    rq_activate_all_grippers(True)
    # end: URCap Program Node
  end
  $ 55 "zero_ftsensor()"
  zero_ftsensor()
  $ 56 "EXTT"
  $ 57 "Set GRP_3F_Enable=Off"
  set_standard_digital_out(4, False)
  $ 58 "Set BarcodeTrigger=Off"
  set_standard_digital_out(6, False)
  $ 59 "Set GRP_3F_Decap=Off"
  set_standard_digital_out(3, False)
  $ 60 "Set GRP_3F_Cap=Off"
  set_standard_digital_out(2, False)
  $ 61 "Set GRP_3F_Open=Off"
  set_standard_digital_out(5, False)
  $ 62 "PSE_T≔get_tool_free_pose(dir=[0,0,0.150], move_in_base_frame=True)"
  global PSE_T=get_tool_free_pose(dir=[0,0,0.150], move_in_base_frame=True)
  $ 63 "If is_reachable(Base_const, [PSE_T])"
  if (is_reachable(p[0.0,0.0,0.0,0.0,0.0,0.0], [PSE_T])):
    $ 64 "MoveL"
    $ 65 "PSE_T" "breakAfter"
    movel(PSE_T, a=1.2, v=0.15)
  end
  while (True):
    $ 66 "Robot Program"
    $ 67 "MAIN"
    $ 68 "command_manager(external_control='uGO', cond_suspend=(ITM_Manipulated and AMR_AtTarget and AMR_Charging and AMR_Battery<40), cond_unsuspend=(AMR_Battery≟60))"
    command_manager(external_control="uGO", cond_suspend=(ITM_Manipulated  and  AMR_AtTarget  and  AMR_Charging  and  AMR_Battery<40), cond_unsuspend=(AMR_Battery == 60))
    $ 69 "log_state(STATE_Info)"
    log_state(STATE_Info)
    $ 70 "Switch STATE"
    switch_1 = STATE
    $ 71 "Case 1"
    if (1 == switch_1):
      $ 72 "Stopping"
      $ 73 "STATE_Info≔'Stopping'"
      global STATE_Info="Stopping"
      $ 74 "end_freedrive_mode()"
      end_freedrive_mode()
      $ 75 "Set"
      set_tcp(p[0.0,0.0,0.161,3.1415,0.0,0.0])
      $ 76 "PSE_T≔get_tool_free_pose(dir=[0,0,0.150], move_in_base_frame=True)"
      global PSE_T=get_tool_free_pose(dir=[0,0,0.150], move_in_base_frame=True)
      $ 77 "If is_reachable(Base_const, [PSE_T])"
      if (is_reachable(p[0.0,0.0,0.0,0.0,0.0,0.0], [PSE_T])):
        $ 78 "MoveL"
        $ 79 "PSE_T" "breakAfter"
        movel(PSE_T, a=1.2, v=0.15)
      end
      $ 80 "do_transition(keep_rxry=OBJ_Picked, r=0)"
      do_transition(keep_rxry=OBJ_Picked, r=0)
      $ 81 "Decapper"
      $ 82 "Set GRP_3F_Enable=Off"
      set_standard_digital_out(4, False)
      $ 83 "Set BarcodeTrigger=Off"
      set_standard_digital_out(6, False)
      $ 84 "Set GRP_3F_Decap=Off"
      set_standard_digital_out(3, False)
      $ 85 "Set GRP_3F_Cap=Off"
      set_standard_digital_out(2, False)
      $ 86 "Set GRP_3F_Open=Off"
      set_standard_digital_out(5, False)
      $ 89 "Call Sub_AMR_MiR_V3"
      Sub_AMR_MiR_V3()
      $ 90 "If stopping() and AMR_Done"
      if (stopping()  and  AMR_Done):
        $ 91 "STATE≔2"
        global STATE=2
        $ 92 "ugo_update_outputs()"
        ugo_update_outputs()
      end
    elif (2 == switch_1):
      $ 93 "Case 2"
      $ 94 "Stopped"
      $ 95 "STATE_Info≔'Stopped'"
      global STATE_Info="Stopped"
      $ 96 "Call Sub_AMR_MiR_V3"
      Sub_AMR_MiR_V3()
      $ 97 "If CMD_Reset"
      if (CMD_Reset):
        $ 98 "STATE≔3"
        global STATE=3
        $ 99 "ugo_update_outputs()"
        ugo_update_outputs()
      end
    elif (3 == switch_1):
      $ 100 "Case 3"
      $ 101 " Resetting"
      $ 102 "STATE_Info≔'Resetting'"
      global STATE_Info="Resetting"
      $ 103 "uML"
      $ 104 "reset_error()"
      reset_error()
      $ 105 "reset_warning()"
      reset_warning()
      $ 106 "PROCESS_Step≔0"
      global PROCESS_Step=0
      $ 107 "PROCESS_Info≔''"
      global PROCESS_Info=""
      $ 108 "ARM_Referenced≔ False "
      global ARM_Referenced=  False
      $ 109 "WRK_Done≔ False "
      global WRK_Done=  False
      $ 110 "ITM_Prepared≔ False "
      global ITM_Prepared=  False
      $ 111 "ITM_Manipulated≔ False "
      global ITM_Manipulated=  False
      $ 112 "STP≔0"
      global STP=0
      $ 113 "Action≔0"
      global Action=0
      $ 114 "Action_Info≔''"
      global Action_Info=""
      $ 115 "ITM_ID≔0"
      global ITM_ID=0
      $ 116 "JIG≔0"
      global JIG=0
      $ 117 "JIG_Slot≔0"
      global JIG_Slot=0
      $ 118 "Task_info≔''"
      global Task_info=""
      $ 119 "Set"
      set_tcp(p[0.0,0.0,0.161,3.1415,0.0,0.0])
      $ 120 "App"
      $ 121 "'ADD APPLICATION SPECIFIC COMMANDS'"
      # 'ADD APPLICATION SPECIFIC COMMANDS'
      $ 122 "OBJ_Type≔0"
      global OBJ_Type=0
      $ 123 "OBJ_Nbr≔0"
      global OBJ_Nbr=0
      $ 124 "If CNT_Rack_Output≥50"
      if (CNT_Rack_Output >= 50):
        $ 125 "CNT_Rack_Output≔0"
        global CNT_Rack_Output=0
      end
      $ 126 "TASK≔struct(ID=0, NAVI=struct(target=0, footprint=0, protectiveOff=0, dock=0), WORK=struct(ITM_ID_Src=0, JIG_ID_Src=0, OBJ_Nbr_Src=0, ACT_Src=0, ITM_ID_Tgt=0, JIG_ID_Tgt=0, OBJ_Nbr_Tgt=0, ACT_Tgt=0, OBJ_Type=0))"
      global TASK=struct(ID=0, NAVI=struct(target=0, footprint=0, protectiveOff=0, dock=0), WORK=struct(ITM_ID_Src=0, JIG_ID_Src=0, OBJ_Nbr_Src=0, ACT_Src=0, ITM_ID_Tgt=0, JIG_ID_Tgt=0, OBJ_Nbr_Tgt=0, ACT_Tgt=0, OBJ_Type=0))
      $ 127 "Call Sub_AMR_MiR_V3"
      Sub_AMR_MiR_V3()
      $ 128 "If resetting() and AMR_Done"
      if (resetting()  and  AMR_Done):
        $ 129 "STATE≔4"
        global STATE=4
        $ 130 "ugo_update_outputs()"
        ugo_update_outputs()
      end
    elif (4 == switch_1):
      $ 131 "Case 4"
      $ 132 "Idle"
      $ 133 "STATE_Info≔'Idle'"
      global STATE_Info="Idle"
      $ 134 "If CMD_Start"
      if (CMD_Start):
        $ 135 "STATE≔5"
        global STATE=5
        $ 136 "ugo_update_outputs()"
        ugo_update_outputs()
      end
    elif (5 == switch_1):
      $ 137 "Case 5"
      $ 138 "Starting"
      $ 139 "STATE_Info≔'Starting'"
      global STATE_Info="Starting"
      $ 140 "'ADD COMMANDS WHAT TO START WITH'"
      # 'ADD COMMANDS WHAT TO START WITH'
      $ 141 "Call Sub_AMR_MiR_V3"
      Sub_AMR_MiR_V3()
      $ 142 "get ugo data"
      $ 143 "Assign Tasks"
      $ 144 "TASK.ID = ugo_get_task()"
      TASK.ID = ugo_get_task()
      $ 145 "If TASK.ID≟1"
      if (TASK.ID == 1):
        $ 146 "Task_info≔'Charge'"
        global Task_info="Charge"
        $ 147 "Parameters"
        $ 148 "AMR_PosTarget≔1"
        global AMR_PosTarget=1
      else:
        $ 149 "ElseIf TASK.ID≟9"
        if (TASK.ID == 9):
          $ 150 "'Pick Sarstedt Rack from Variable source'"
          # 'Pick Sarstedt Rack from Variable source'
          $ 151 "Task_info≔'Navigate to Target'"
          global Task_info="Navigate to Target"
          $ 152 "Parameters"
          $ 153 "AMR_PosTarget≔UGO.read_input('00','ITM_ID')"
          global AMR_PosTarget=UGO.read_input("00","ITM_ID")
        else:
          $ 154 "ElseIf TASK.ID≟10"
          if (TASK.ID == 10):
            $ 155 "'Pick Sarstedt Rack from Variable source'"
            # 'Pick Sarstedt Rack from Variable source'
            $ 156 "Task_info≔'Pick Rack'"
            global Task_info="Pick Rack"
            $ 157 "AMR_PosTarget≔2"
            global AMR_PosTarget=2
            $ 158 "Parameters"
            $ 159 "ITM_ID≔UGO.read_input('00','ITM_ID')"
            global ITM_ID=UGO.read_input("00","ITM_ID")
            $ 160 "JIG≔UGO.read_input('00','JIG_ID')"
            global JIG=UGO.read_input("00","JIG_ID")
            $ 161 "OBJ_Type≔3"
            global OBJ_Type=3
          else:
            $ 163 "ElseIf TASK.ID≟11"
            if (TASK.ID == 11):
              $ 164 "'Place Sarstedt Rack on Variable target'"
              # 'Place Sarstedt Rack on Variable target'
              $ 165 "Task_info≔'Place Rack'"
              global Task_info="Place Rack"
              $ 166 "AMR_PosTarget≔2"
              global AMR_PosTarget=2
              $ 167 "Parameters"
              $ 168 "ITM_ID≔UGO.read_input('00','ITM_ID')"
              global ITM_ID=UGO.read_input("00","ITM_ID")
              $ 169 "JIG≔UGO.read_input('00','JIG_ID')"
              global JIG=UGO.read_input("00","JIG_ID")
              $ 170 "OBJ_Type≔3"
              global OBJ_Type=3
            else:
              $ 172 "ElseIf TASK.ID≟12"
              if (TASK.ID == 12):
                $ 173 "Task_info≔'Decapping'"
                global Task_info="Decapping"
                $ 174 "Parameters"
                $ 175 "ITM_ID≔1"
                global ITM_ID=1
                $ 176 "AMR_PosTarget≔AMR_PosActual"
                global AMR_PosTarget=AMR_PosActual
                $ 177 "PRC_TubCounter≔0"
                global PRC_TubCounter=0
              else:
                $ 178 "ElseIf TASK.ID≟13"
                if (TASK.ID == 13):
                  $ 179 "Task_info≔'Empty racks'"
                  global Task_info="Empty racks"
                  $ 180 "Parameters"
                  $ 181 "ITM_ID≔1"
                  global ITM_ID=1
                  $ 182 "AMR_PosTarget≔AMR_PosActual"
                  global AMR_PosTarget=AMR_PosActual
                else:
                  $ 183 "ElseIf TASK.ID≟14"
                  if (TASK.ID == 14):
                    $ 184 "Task_info≔'Decap'"
                    global Task_info="Decap"
                    $ 185 "Parameters"
                    $ 186 "ITM_ID≔1"
                    global ITM_ID=1
                    $ 187 "OBJ_Type≔2"
                    global OBJ_Type=2
                    $ 188 "JIG≔7"
                    global JIG=7
                    $ 189 "AMR_PosTarget≔AMR_PosActual"
                    global AMR_PosTarget=AMR_PosActual
                  else:
                    $ 190 "ElseIf TASK.ID≟99"
                    if (TASK.ID == 99):
                      $ 191 "Task_info≔'Decapping and barcode alignment'"
                      global Task_info="Decapping and barcode alignment"
                      $ 192 "Parameters"
                      $ 193 "PRC_TubNumber≔UGO.read_input('00','TubesNb')"
                      global PRC_TubNumber=UGO.read_input("00","TubesNb")
                      $ 194 "PRC_TubCounter≔0"
                      global PRC_TubCounter=0
                      $ 195 "ITM_ID≔1"
                      global ITM_ID=1
                      $ 196 "AMR_PosTarget≔AMR_PosActual"
                      global AMR_PosTarget=AMR_PosActual
                    else:
                      $ 205 "ElseIf TASK.ID≟15"
                      if (TASK.ID == 15):
                        $ 206 "Task_info≔'Unoad Centrifuge'"
                        global Task_info="Unoad Centrifuge"
                        $ 207 "Parameters"
                        $ 208 "PRC_RackCounter≔0"
                        global PRC_RackCounter=0
                        $ 209 "TASK.WORK.ITM_ID_Src=2"
                        TASK.WORK.ITM_ID_Src=2
                        $ 210 "TASK.WORK.ITM_ID_Tgt=1"
                        TASK.WORK.ITM_ID_Tgt=1
                        $ 211 "AMR_PosTarget≔4"
                        global AMR_PosTarget=4
                        $ 212 "AMR_FootprintID≔1"
                        global AMR_FootprintID=1
                      else:
                        $ 231 "Else" "noBreak"
                        $ 232 "set_error(ERROR_WRONG_ORDER)"
                        set_error(ERROR_WRONG_ORDER)
                      end
                    end
                  end
                end
              end
            end
          end
        end
      end
      $ 233 "test ugo"
      $ 234 "Wait: 0.2"
      sleep(0.2)
      $ 235 "ugo_update_outputs()"
      ugo_update_outputs()
      $ 236 "If starting() and AMR_Done"
      if (starting()  and  AMR_Done):
        $ 237 "log_message(Task_info, 'New Task: ')"
        log_message(Task_info, "New Task: ")
        $ 238 "log_message(to_str(TASK.ID), 'Task_ID: ')"
        log_message(to_str(TASK.ID), "Task_ID: ")
        $ 239 "do_transition(keep_rxry=OBJ_Picked)"
        do_transition(keep_rxry=OBJ_Picked)
        $ 240 "STATE≔6"
        global STATE=6
        $ 241 "ugo_update_outputs()"
        ugo_update_outputs()
      end
    elif (6 == switch_1):
      $ 242 "Case 6"
      $ 243 "Execute"
      $ 244 "STATE_Info≔'Execute'"
      global STATE_Info="Execute"
      $ 245 "If  not CMD_Hold and not CMD_Suspend"
      global thread_flag_245=0
      thread Thread_if_245():
        $ 246 "Switch PROCESS_Step"
        switch_2 = PROCESS_Step
        $ 247 "Case 0"
        if (0 == switch_2):
          $ 248 "PROCESS_Info≔'process control'"
          global PROCESS_Info="process control"
          $ 249 "log_process(PROCESS_Info)"
          log_process(PROCESS_Info)
          $ 250 "process control"
          $ 251 "If  not AMR_AtTarget"
          if (  not  AMR_AtTarget):
            $ 252 "PROCESS_Step≔1"
            global PROCESS_Step=1
          else:
            $ 253 "ElseIf (( not ITM_Prepared and  not WRK_Done) or (ITM_Prepared and WRK_Done))"
            if (((  not  ITM_Prepared  and    not  WRK_Done)  or  (ITM_Prepared  and  WRK_Done))):
              $ 254 "PROCESS_Step≔2"
              global PROCESS_Step=2
            else:
              $ 255 "ElseIf  not WRK_Done"
              if (  not  WRK_Done):
                $ 256 "PROCESS_Step≔3"
                global PROCESS_Step=3
              else:
                $ 257 "Else" "noBreak"
                $ 258 "task finished"
                $ 259 "PROCESS_Info≔''"
                global PROCESS_Info=""
                $ 260 "STATE≔7"
                global STATE=7
                $ 261 "ugo_update_outputs()"
                ugo_update_outputs()
              end
            end
          end
        elif (1 == switch_2):
          $ 262 "Case 1"
          $ 263 "navigate"
          $ 264 "'MOVING THE uML'"
          # 'MOVING THE uML'
          $ 265 "PROCESS_Info≔'move to target'"
          global PROCESS_Info="move to target"
          $ 266 "log_process(PROCESS_Info)"
          log_process(PROCESS_Info)
          $ 267 "If TASK.ID≟1"
          if (TASK.ID == 1):
            $ 268 "Action≔51"
            global Action=51
          else:
            $ 269 "Else" "noBreak"
            $ 270 "Action≔52"
            global Action=52
          end
          $ 271 "Call Sub_AMR_MiR_V3"
          Sub_AMR_MiR_V3()
          $ 272 "If AMR_Done"
          if (AMR_Done):
            $ 273 "PROCESS_Step≔0"
            global PROCESS_Step=0
          end
        elif (2 == switch_2):
          $ 274 "Case 2"
          $ 275 "prepare"
          $ 276 "'THINGS THAT HAVE TO BE DONE ONCE IN A SEQUENCE,WORKFLOW'"
          # 'THINGS THAT HAVE TO BE DONE ONCE IN A SEQUENCE,WORKFLOW'
          $ 277 "PROCESS_Info≔'prepare for work'"
          global PROCESS_Info="prepare for work"
          $ 278 "log_process(PROCESS_Info)"
          log_process(PROCESS_Info)
          $ 279 "If TASK.WORK.ITM_ID_Src>1"
          if (TASK.WORK.ITM_ID_Src>1):
            $ 280 "ITM_ID≔TASK.WORK.ITM_ID_Src"
            global ITM_ID=TASK.WORK.ITM_ID_Src
          else:
            $ 281 "ElseIf TASK.WORK.ITM_ID_Tgt>1"
            if (TASK.WORK.ITM_ID_Tgt>1):
              $ 282 "ITM_ID≔TASK.WORK.ITM_ID_Tgt"
              global ITM_ID=TASK.WORK.ITM_ID_Tgt
            end
          end
          $ 283 "If  not ARM_Referenced and (ITM_ID≠0)"
          if (  not  ARM_Referenced  and  (ITM_ID != 0)):
            $ 284 "STP≔1"
            global STP=1
          else:
            $ 285 "ElseIf ARM_Referenced or (ITM_ID≟0)"
            if (ARM_Referenced  or  (ITM_ID == 0)):
              $ 286 "STP≔2"
              global STP=2
            end
          end
          $ 287 "Switch STP"
          switch_3 = STP
          $ 288 "Case 1"
          if (1 == switch_3):
            $ 289 "reference"
            $ 290 "STP_Info≔'reference at target position'"
            global STP_Info="reference at target position"
            $ 291 "log_step(STP_Info)"
            log_step(STP_Info)
            $ 292 "If ITM_ID≟1"
            if (ITM_ID == 1):
              $ 293 "CAM_Done≔ True "
              global CAM_Done=  True
            else:
              $ 294 "Else" "noBreak"
              $ 295 "Action≔131"
              global Action=131
              $ 296 "Call Sub_Vision_V18"
              Sub_Vision_V18()
            end
            $ 298 "If CAM_Done and  not ERROR.FLAG"
            if (CAM_Done  and    not  ERROR.FLAG):
              $ 299 "log_step('ARM referenced')"
              log_step("ARM referenced")
              $ 300 "ARM_Referenced≔ True "
              global ARM_Referenced=  True
            end
          elif (2 == switch_3):
            $ 301 "Case 2"
            $ 302 "manipulate"
            $ 303 "STP_Info≔'manipulate item'"
            global STP_Info="manipulate item"
            $ 304 "log_step(STP_Info)"
            log_step(STP_Info)
            $ 305 "'In case pressing button is needed'"
            # 'In case pressing button is needed'
            $ 306 "If found_in_list(ITM_ID, ITM_ID_List)"
            if (found_in_list(ITM_ID, ITM_ID_List)):
              $ 307 "Switch ITM_ID"
              switch_4 = ITM_ID
              $ 308 "Case 0"
              if (0 == switch_4):
                $ 309 "ITM_Manipulated≔ not ITM_Manipulated"
                global ITM_Manipulated=  not  ITM_Manipulated
              elif (1 == switch_4):
                $ 310 "Case 1"
                $ 311 "ITM_Manipulated≔ not ITM_Manipulated"
                global ITM_Manipulated=  not  ITM_Manipulated
              elif (2 == switch_4):
                $ 312 "Case 2"
              else:
                $ 322 "Default Case"
                $ 323 "ITM_Manipulated≔ not ITM_Manipulated"
                global ITM_Manipulated=  not  ITM_Manipulated
              end
            end
          end
          $ 324 "ITM_Prepared≔(ITM_Manipulated or  not found_in_list(ITM_ID, ITM_ID_List)) and (ARM_Referenced or ITM_ID≟0) and  not WRK_Done"
          global ITM_Prepared=(ITM_Manipulated  or    not  found_in_list(ITM_ID, ITM_ID_List))  and  (ARM_Referenced  or  ITM_ID == 0)  and    not  WRK_Done
          $ 325 "STP≔0"
          global STP=0
          $ 326 "STP_Info≔''"
          global STP_Info=""
          $ 327 "PROCESS_Step≔0"
          global PROCESS_Step=0
        elif (3 == switch_2):
          $ 328 "Case 3"
          $ 329 "work"
          $ 330 "'ADD EVERY MACHINE, OBJECT, STATION TO WORK ON'"
          # 'ADD EVERY MACHINE, OBJECT, STATION TO WORK ON'
          $ 331 "Switch ITM_ID"
          switch_3 = ITM_ID
          $ 332 "Case 1"
          if (1 == switch_3):
            $ 333 "uLM"
            $ 334 "If TASK.ID≟12"
            if (TASK.ID == 12):
              $ 335 "fill racks"
              $ 336 "Action≔151"
              global Action=151
              $ 337 "Call Sub_Vision_V18"
              Sub_Vision_V18()
              $ 338 "If  not ERROR.FLAG"
              if (  not  ERROR.FLAG):
                $ 339 "Actions for the task"
                $ 340 "Action≔1"
                global Action=1
                $ 341 "JIG≔2"
                global JIG=2
                $ 342 "JIG_Slot≔CAM_Result[0]"
                global JIG_Slot=CAM_Result[0]
                $ 343 "OBJ_Nbr≔CAM_Result[0]"
                global OBJ_Nbr=CAM_Result[0]
                $ 344 "OBJ_Type≔2"
                global OBJ_Type=2
                $ 345 "Call Sub_Action_V4"
                Sub_Action_V4()
                $ 346 "If OBJ_Picked"
                if (OBJ_Picked):
                  $ 347 "CAM_Result.remove(0)"
                  CAM_Result.remove(0)
                  $ 348 "PRC_TubCounter≔PRC_TubCounter+1"
                  global PRC_TubCounter=PRC_TubCounter+1
                  $ 349 "If PRC_TubCounter%4≟0"
                  if (PRC_TubCounter%4 == 0):
                    $ 350 "JIG_Slot≔4"
                    global JIG_Slot=4
                  else:
                    $ 351 "Else" "noBreak"
                    $ 352 "JIG_Slot≔PRC_TubCounter%4"
                    global JIG_Slot=PRC_TubCounter%4
                  end
                  $ 353 "OBJ_Nbr≔ceil(PRC_TubCounter/4)"
                  global OBJ_Nbr=ceil(PRC_TubCounter/4)
                  $ 354 "Action≔2"
                  global Action=2
                  $ 355 "JIG≔4"
                  global JIG=4
                  $ 356 "Call Sub_Action_V4"
                  Sub_Action_V4()
                  $ 357 "Action≔151"
                  global Action=151
                  $ 358 "Call Sub_Vision_V18"
                  Sub_Vision_V18()
                end
              end
              $ 359 "If (CAM_Captures≥CAM_PRM_Retries) or (PRC_TubCounter≥32)"
              if ((CAM_Captures >= CAM_PRM_Retries)  or  (PRC_TubCounter >= 32)):
                $ 360 "PROCESS_Step≔0"
                global PROCESS_Step=0
                $ 361 "WRK_Done≔ True "
                global WRK_Done=  True
              end
            else:
              $ 362 "ElseIf TASK.ID≟10"
              if (TASK.ID == 10):
                $ 363 "Pick Rack"
                $ 364 "Action≔131"
                global Action=131
                $ 365 "Call Sub_Vision_V18"
                Sub_Vision_V18()
                $ 366 "Action≔1"
                global Action=1
                $ 367 "Call Sub_Action_V4"
                Sub_Action_V4()
                $ 368 "PROCESS_Step≔0"
                global PROCESS_Step=0
                $ 369 "WRK_Done≔ True "
                global WRK_Done=  True
              else:
                $ 370 "ElseIf TASK.ID≟11"
                if (TASK.ID == 11):
                  $ 371 "Place Rack"
                  $ 372 "Action≔2"
                  global Action=2
                  $ 373 "Call Sub_Action_V4"
                  Sub_Action_V4()
                  $ 374 "PROCESS_Step≔0"
                  global PROCESS_Step=0
                  $ 375 "WRK_Done≔ True "
                  global WRK_Done=  True
                else:
                  $ 376 "ElseIf TASK.ID≟13"
                  if (TASK.ID == 13):
                    $ 377 "empty racks"
                    $ 378 "pick"
                    $ 379 "Action≔1"
                    global Action=1
                    $ 380 "JIG≔4"
                    global JIG=4
                    $ 381 "If PRC_TubCounter%4≟0"
                    if (PRC_TubCounter%4 == 0):
                      $ 382 "JIG_Slot≔4"
                      global JIG_Slot=4
                    else:
                      $ 383 "Else" "noBreak"
                      $ 384 "JIG_Slot≔PRC_TubCounter%4"
                      global JIG_Slot=PRC_TubCounter%4
                    end
                    $ 385 "OBJ_Nbr≔ceil(PRC_TubCounter/4)"
                    global OBJ_Nbr=ceil(PRC_TubCounter/4)
                    $ 386 "OBJ_Type≔2"
                    global OBJ_Type=2
                    $ 387 "Call Sub_Action_V4"
                    Sub_Action_V4()
                    $ 388 "If OBJ_Picked"
                    if (OBJ_Picked):
                      $ 389 "Action≔2"
                      global Action=2
                      $ 390 "JIG≔3"
                      global JIG=3
                      $ 391 "JIG_Slot≔1"
                      global JIG_Slot=1
                      $ 392 "CNT_Rack_Output≔CNT_Rack_Output + 1"
                      global CNT_Rack_Output=CNT_Rack_Output + 1
                      $ 393 "OBJ_Nbr≔CNT_Rack_Output"
                      global OBJ_Nbr=CNT_Rack_Output
                      $ 394 "Call Sub_Action_V4"
                      Sub_Action_V4()
                      $ 395 "If  not ERROR.FLAG"
                      if (  not  ERROR.FLAG):
                        $ 396 "PRC_TubCounter≔PRC_TubCounter - 1"
                        global PRC_TubCounter=PRC_TubCounter - 1
                      end
                    end
                    $ 397 "If CNT_Rack_Output≥50 or PRC_TubCounter≤0"
                    if (CNT_Rack_Output >= 50  or  PRC_TubCounter <= 0):
                      $ 398 "PROCESS_Step≔0"
                      global PROCESS_Step=0
                      $ 399 "WRK_Done≔ True "
                      global WRK_Done=  True
                    end
                  else:
                    $ 400 "ElseIf TASK.ID≟14"
                    if (TASK.ID == 14):
                      $ 403 "samples≔ True "
                      global samples=  True
                      $ 404 "Loop samples≟ True "
                      while (samples ==   True  ):
                        $ 405 "JIG≔7"
                        global JIG=7
                        $ 406 "Action≔151"
                        global Action=151
                        $ 407 "Call Sub_Vision_V18"
                        Sub_Vision_V18()
                        $ 408 "Action≔1"
                        global Action=1
                        $ 409 "JIG≔2"
                        global JIG=2
                        $ 410 "JIG_Slot≔CAM_Result[0]"
                        global JIG_Slot=CAM_Result[0]
                        $ 411 "OBJ_Nbr≔CAM_Result[0]"
                        global OBJ_Nbr=CAM_Result[0]
                        $ 412 "OBJ_Type≔2"
                        global OBJ_Type=2
                        $ 413 "Call Sub_Action_V4"
                        Sub_Action_V4()
                        $ 414 "JIG≔1"
                        global JIG=1
                        $ 415 "Action≔11"
                        global Action=11
                        $ 416 "Call Sub_Action_V4"
                        Sub_Action_V4()
                        $ 417 "Action≔12"
                        global Action=12
                        $ 418 "Call Sub_Action_V4"
                        Sub_Action_V4()
                        $ 419 "Action≔2"
                        global Action=2
                        $ 420 "JIG≔6"
                        global JIG=6
                        $ 421 "Call Sub_Action_V4"
                        Sub_Action_V4()
                        $ 422 "Action≔13"
                        global Action=13
                        $ 423 "Call Sub_Action_V4"
                        Sub_Action_V4()
                        $ 424 "Action≔1"
                        global Action=1
                        $ 425 "JIG≔1"
                        global JIG=1
                        $ 426 "Call Sub_Action_V4"
                        Sub_Action_V4()
                        $ 427 "JIG≔2"
                        global JIG=2
                        $ 428 "Action≔2"
                        global Action=2
                        $ 431 "OBJ_Type≔2"
                        global OBJ_Type=2
                        $ 432 "Call Sub_Action_V4"
                        Sub_Action_V4()
                      end
                    end
                  end
                end
              end
            end
          elif (2 == switch_3):
            $ 433 "Case 2"
          elif (20 == switch_3):
            $ 475 "Case 20"
          else:
            $ 537 "Default Case"
            $ 538 "WRK_Done≔ True "
            global WRK_Done=  True
            $ 539 "PROCESS_Step≔0"
            global PROCESS_Step=0
          end
        end
        thread_flag_245 = 1
      end
      if (  not  CMD_Hold and not CMD_Suspend):
        global thread_handler_245=run Thread_if_245()
        while (thread_flag_245 == 0):
          if not(  not  CMD_Hold and not CMD_Suspend):
            kill thread_handler_245
            thread_flag_245 = 2
          else:
            sync()
          end
        end
      else:
        thread_flag_245 = 2
      end
      $ 540 "If CMD_Hold"
      if (CMD_Hold):
        $ 541 "STATE≔9"
        global STATE=9
        $ 542 "ugo_update_outputs()"
        ugo_update_outputs()
      else:
        $ 543 "ElseIf CMD_Suspend"
        if (CMD_Suspend):
          $ 544 "STATE≔12"
          global STATE=12
          $ 545 "ugo_update_outputs()"
          ugo_update_outputs()
        end
      end
    elif (7 == switch_1):
      $ 546 "Case 7"
      $ 547 "Completing"
      $ 548 "STATE_Info≔'Completing'"
      global STATE_Info="Completing"
      $ 549 "'ADD COMMANDS FOR COMPLETING THE PROCESS'"
      # 'ADD COMMANDS FOR COMPLETING THE PROCESS'
      $ 550 "do_transition(keep_rxry=OBJ_Picked)"
      do_transition(keep_rxry=OBJ_Picked)
      $ 551 "Call Sub_AMR_MiR_V3"
      Sub_AMR_MiR_V3()
      $ 552 "If completing() and AMR_Done"
      if (completing()  and  AMR_Done):
        $ 553 "STATE≔8"
        global STATE=8
        $ 554 "ugo_update_outputs()"
        ugo_update_outputs()
      end
    elif (8 == switch_1):
      $ 555 "Case 8"
      $ 556 "Complete"
      $ 557 "STATE_Info≔'Complete'"
      global STATE_Info="Complete"
      $ 558 "If CMD_Reset"
      if (CMD_Reset):
        $ 559 "STATE≔3"
        global STATE=3
        $ 560 "ugo_update_outputs()"
        ugo_update_outputs()
      end
    elif (9 == switch_1):
      $ 561 "Case 9"
      $ 562 "Holding"
      $ 563 "STATE_Info≔'Holding'"
      global STATE_Info="Holding"
      $ 564 "stopl(0.5)"
      stopl(0.5)
      $ 565 "Call Sub_AMR_MiR_V3"
      Sub_AMR_MiR_V3()
      $ 566 "If holding() and AMR_Done"
      if (holding()  and  AMR_Done):
        $ 567 "STATE≔10"
        global STATE=10
        $ 568 "ugo_update_outputs()"
        ugo_update_outputs()
      end
    elif (10 == switch_1):
      $ 569 "Case 10"
      $ 570 "Held"
      $ 571 "STATE_Info≔'Held'"
      global STATE_Info="Held"
      $ 572 "If CMD_Unhold"
      if (CMD_Unhold):
        $ 573 "end_freedrive_mode()"
        end_freedrive_mode()
        $ 574 "STATE≔11"
        global STATE=11
        $ 575 "ugo_update_outputs()"
        ugo_update_outputs()
      else:
        $ 576 "ElseIf FNC_Freedrive"
        if (FNC_Freedrive):
          $ 577 "freedrive_mode()"
          freedrive_mode()
        else:
          $ 578 "Else" "noBreak"
          $ 579 "end_freedrive_mode()"
          end_freedrive_mode()
        end
      end
    elif (11 == switch_1):
      $ 580 "Case 11"
      $ 581 "Unholding"
      $ 582 "STATE_Info≔'Unholding'"
      global STATE_Info="Unholding"
      $ 583 "Clearing"
      $ 584 "Switch ERROR.ID"
      switch_2 = ERROR.ID
      $ 585 "Case 1002"
      if (1002 == switch_2):
        $ 586 "AMR_AtTarget≔ False "
        global AMR_AtTarget=  False
        $ 587 "ARM_Referenced≔ False "
        global ARM_Referenced=  False
        $ 588 "ITM_Prepared≔ False "
        global ITM_Prepared=  False
        $ 589 "PROCESS_Step≔1"
        global PROCESS_Step=1
      elif (2007 == switch_2):
        $ 590 "Case 2007"
        $ 591 "PROCESS_Step≔1"
        global PROCESS_Step=1
      end
      $ 592 "reset_error()"
      reset_error()
      $ 593 "reset_warning()"
      reset_warning()
      $ 594 "OBJ_Picked≔gripper_has_object()"
      global OBJ_Picked=gripper_has_object()
      $ 595 "Call Sub_AMR_MiR_V3"
      Sub_AMR_MiR_V3()
      $ 596 "If unholding() and AMR_Done"
      if (unholding()  and  AMR_Done):
        $ 597 "STATE≔6"
        global STATE=6
        $ 598 "ugo_update_outputs()"
        ugo_update_outputs()
      end
    elif (12 == switch_1):
      $ 599 "Case 12"
      $ 600 "Suspending"
      $ 601 "STATE_Info≔'Suspending'"
      global STATE_Info="Suspending"
      $ 602 "PROCESS_Info≔str_cat(PROCESS_Info, ' suspended')"
      global PROCESS_Info=str_cat(PROCESS_Info, " suspended")
      $ 603 "If suspending()"
      if (suspending()):
        $ 604 "STATE≔13"
        global STATE=13
        $ 605 "ugo_update_outputs()"
        ugo_update_outputs()
      end
    elif (13 == switch_1):
      $ 606 "Case 13"
      $ 607 "Suspended"
      $ 608 "STATE_Info≔'Suspended'"
      global STATE_Info="Suspended"
      $ 609 "Call Sub_AMR_MiR_V3"
      Sub_AMR_MiR_V3()
      $ 610 "If CMD_Unsuspend"
      if (CMD_Unsuspend):
        $ 611 "STATE≔14"
        global STATE=14
        $ 612 "ugo_update_outputs()"
        ugo_update_outputs()
      end
    elif (14 == switch_1):
      $ 613 "Case 14"
      $ 614 "Unsuspending"
      $ 615 "STATE_Info≔'Unsuspending'"
      global STATE_Info="Unsuspending"
      $ 616 "PROCESS_Step≔0"
      global PROCESS_Step=0
      $ 617 "If unsuspending()"
      if (unsuspending()):
        $ 618 "STATE≔6"
        global STATE=6
        $ 619 "ugo_update_outputs()"
        ugo_update_outputs()
      end
    elif (15 == switch_1):
      $ 620 "Case 15"
      $ 621 "Aborting"
      $ 622 "STATE_Info≔'Aborting'"
      global STATE_Info="Aborting"
      $ 623 "If aborting()"
      if (aborting()):
        $ 624 "STATE≔16"
        global STATE=16
        $ 625 "ugo_update_outputs()"
        ugo_update_outputs()
      end
    elif (16 == switch_1):
      $ 626 "Case 16"
      $ 627 "Aborted"
      $ 628 "STATE_Info≔'Aborted'"
      global STATE_Info="Aborted"
      $ 629 "If CMD_Clear"
      if (CMD_Clear):
        $ 630 "STATE≔17"
        global STATE=17
        $ 631 "ugo_update_outputs()"
        ugo_update_outputs()
      end
    elif (17 == switch_1):
      $ 632 "Case 17"
      $ 633 "Clearing"
      $ 634 "STATE_Info≔'Clearing'"
      global STATE_Info="Clearing"
      $ 635 "Clearing"
      $ 636 "reset_warning()"
      reset_warning()
      $ 637 "reset_error()"
      reset_error()
      $ 638 "If clearing()"
      if (clearing()):
        $ 639 "STATE≔2"
        global STATE=2
        $ 640 "ugo_update_outputs()"
        ugo_update_outputs()
      end
    end
    $ 641 "log_state(STATE_Info)"
    log_state(STATE_Info)
    $ 642 "log_warning(WARNING.MSG)"
    log_warning(WARNING.MSG)
    $ 643 "log_error(ERROR.MSG)"
    log_error(ERROR.MSG)
    $ 644 "Times"
    $ 645 "Switch STATE"
    switch_1 = STATE
    $ 646 "Case 1"
    if (1 == switch_1):
      $ 647 "TM_St_Stopping≔get_time(STATE_Times[STATE-1])"
      global TM_St_Stopping=get_time(STATE_Times[STATE-1])
    elif (2 == switch_1):
      $ 648 "Case 2"
      $ 649 "TM_St_Stopped≔get_time(STATE_Times[STATE-1])"
      global TM_St_Stopped=get_time(STATE_Times[STATE-1])
    elif (3 == switch_1):
      $ 650 "Case 3"
      $ 651 "TM_St_Resetting≔get_time(STATE_Times[STATE-1])"
      global TM_St_Resetting=get_time(STATE_Times[STATE-1])
    elif (4 == switch_1):
      $ 652 "Case 4"
      $ 653 "TM_St_Idle≔get_time(STATE_Times[STATE-1])"
      global TM_St_Idle=get_time(STATE_Times[STATE-1])
    elif (5 == switch_1):
      $ 654 "Case 5"
      $ 655 "TM_St_Starting≔get_time(STATE_Times[STATE-1])"
      global TM_St_Starting=get_time(STATE_Times[STATE-1])
    elif (6 == switch_1):
      $ 656 "Case 6"
      $ 657 "TM_St_Execute≔get_time(STATE_Times[STATE-1])"
      global TM_St_Execute=get_time(STATE_Times[STATE-1])
    elif (7 == switch_1):
      $ 658 "Case 7"
      $ 659 "TM_St_Completin≔get_time(STATE_Times[STATE-1])"
      global TM_St_Completin=get_time(STATE_Times[STATE-1])
    elif (8 == switch_1):
      $ 660 "Case 8"
      $ 661 "TM_St_Complete≔get_time(STATE_Times[STATE-1])"
      global TM_St_Complete=get_time(STATE_Times[STATE-1])
    elif (9 == switch_1):
      $ 662 "Case 9"
      $ 663 "TM_St_Holding≔get_time(STATE_Times[STATE-1])"
      global TM_St_Holding=get_time(STATE_Times[STATE-1])
    elif (10 == switch_1):
      $ 664 "Case 10"
      $ 665 "TM_St_Held≔get_time(STATE_Times[STATE-1])"
      global TM_St_Held=get_time(STATE_Times[STATE-1])
    elif (11 == switch_1):
      $ 666 "Case 11"
      $ 667 "TM_St_Unholding≔get_time(STATE_Times[STATE-1])"
      global TM_St_Unholding=get_time(STATE_Times[STATE-1])
    elif (12 == switch_1):
      $ 668 "Case 12"
      $ 669 "TM_St_Suspendin≔get_time(STATE_Times[STATE-1])"
      global TM_St_Suspendin=get_time(STATE_Times[STATE-1])
    elif (13 == switch_1):
      $ 670 "Case 13"
      $ 671 "TM_St_Suspended≔get_time(STATE_Times[STATE-1])"
      global TM_St_Suspended=get_time(STATE_Times[STATE-1])
    elif (14 == switch_1):
      $ 672 "Case 14"
      $ 673 "TM_St_Unsuspend≔get_time(STATE_Times[STATE-1])"
      global TM_St_Unsuspend=get_time(STATE_Times[STATE-1])
    elif (15 == switch_1):
      $ 674 "Case 15"
      $ 675 "TM_St_Aborting≔get_time(STATE_Times[STATE-1])"
      global TM_St_Aborting=get_time(STATE_Times[STATE-1])
    elif (16 == switch_1):
      $ 676 "Case 16"
      $ 677 "TM_St_Aborted≔get_time(STATE_Times[STATE-1])"
      global TM_St_Aborted=get_time(STATE_Times[STATE-1])
    elif (17 == switch_1):
      $ 678 "Case 17"
      $ 679 "TM_St_Clearing≔get_time(STATE_Times[STATE-1])"
      global TM_St_Clearing=get_time(STATE_Times[STATE-1])
    end
    $ 681 "Wait: 0.1"
    sleep(0.1)
  end
end
